FUNCTION_BLOCK ManualOperation (* Basic Function Block Type *)
  (* Standard: 61499-2 *)
  (* Version 0.0, 10/19/2026, macie, Schneider Electric, Template *)
  PACKAGE Main;
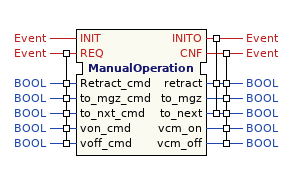
  EVENT_INPUT
    INIT; (* Initialization Request *)
    REQ WITH Retract_cmd, to_mgz_cmd, to_nxt_cmd, von_cmd, voff_cmd; (* Normal Execution Request *)
  END_EVENT
  EVENT_OUTPUT
    INITO WITH retract, to_next; (* Initialization Confirm *)
    CNF WITH retract, to_mgz, to_next, vcm_off, vcm_on; (* Execution Confirmation *)
  END_EVENT
  VAR_INPUT
    Retract_cmd : BOOL; (* Input event qualifier *)
    to_mgz_cmd : BOOL;
    to_nxt_cmd : BOOL;
    von_cmd : BOOL;
    voff_cmd : BOOL;
  END_VAR
  VAR_OUTPUT
    retract : BOOL; (* Output event qualifier *)
    to_mgz : BOOL;
    to_next : BOOL;
    vcm_on : BOOL;
    vcm_off : BOOL;
  END_VAR
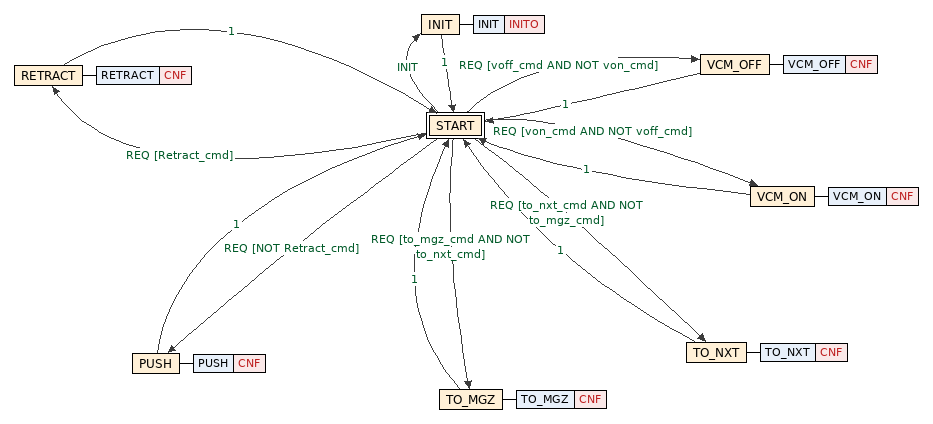
  EC_STATES
    START; (* Initial State *)
    INIT : INIT -> INITO; (* Initialization *)
    RETRACT : RETRACT -> CNF; (* Normal execution *)
    PUSH : PUSH -> CNF;
    TO_MGZ : TO_MGZ -> CNF;
    TO_NXT : TO_NXT -> CNF;
    VCM_ON : VCM_ON -> CNF;
    VCM_OFF : VCM_OFF -> CNF;
  END_STATES
  EC_TRANSITIONS
    START TO INIT := INIT;
    INIT TO START := 1;
    START TO RETRACT := REQ [Retract_cmd];
    RETRACT TO START := 1;
    START TO PUSH := REQ [NOT Retract_cmd];
    PUSH TO START := 1;
    START TO TO_MGZ := REQ [to_mgz_cmd AND NOT to_nxt_cmd];
    TO_MGZ TO START := 1;
    START TO TO_NXT := REQ [to_nxt_cmd AND NOT to_mgz_cmd];
    TO_NXT TO START := 1;
    START TO VCM_ON := REQ [von_cmd AND NOT voff_cmd];
    VCM_ON TO START := 1;
    START TO VCM_OFF := REQ [voff_cmd AND NOT von_cmd];
    VCM_OFF TO START := 1;
  END_TRANSITIONS
  ALGORITHM INIT IN ST: (* Initialization algorithm *)
;
retract := FALSE;
to_mgz := FALSE;
to_next := TRUE;
vcm_off := FALSE;
vcm_on := FALSE;
  END_ALGORITHM
  ALGORITHM RETRACT IN ST: (* Normally executed algorithm *)
;
retract := TRUE;
  END_ALGORITHM
  ALGORITHM PUSH IN ST:
;
retract := FALSE;
  END_ALGORITHM
  ALGORITHM TO_MGZ IN ST:
;
to_mgz := TRUE;
to_next := FALSE;
  END_ALGORITHM
  ALGORITHM TO_NXT IN ST:
;
to_mgz := FALSE;
to_next := TRUE;
  END_ALGORITHM
  ALGORITHM VCM_ON IN ST:
;
vcm_on := TRUE;
vcm_off := FALSE;
  END_ALGORITHM
  ALGORITHM VCM_OFF IN ST:
;

vcm_on := FALSE;
vcm_off := TRUE;
  END_ALGORITHM
END_FUNCTION_BLOCK
